(* IEC 61131-3 sources: plc-vscode/tests/st/all/trust-platform/examples/communication/opcua/src, 2 files *)

(* ---- config.st ---- *)
CONFIGURATION Config
VAR_GLOBAL
    TankLevel : REAL := 42.5;
    PumpRunning : BOOL := FALSE;
END_VAR
RESOURCE CommRes ON PLC
    TASK MainTask (INTERVAL := T#100ms, PRIORITY := 1);
    PROGRAM Main WITH MainTask : Main;
END_RESOURCE
END_CONFIGURATION

(* ---- main.st ---- *)
PROGRAM Main
VAR_EXTERNAL
    TankLevel : REAL;
    PumpRunning : BOOL;
END_VAR

PumpRunning := TankLevel > 50.0;
END_PROGRAM
